(* IEC 61131-3 sources: codesys-api/examples/mqtt_large_payload/st/sfw, 5 files *)

(* ---- FB_MixedPushStream.st ---- *)
FUNCTION_BLOCK FB_MixedPushStream
// One periodic stream of the mixed-rate test through MQTT.MqttStoreForward (MixedPushTest, mixed_rate_test.py --push).
// FB_MixedStream's messages, built the same way (same tags, values, "MIX:<StreamId>:<round>:<part>:<parts>:<UTC ms>"
// header and "<tag>:<value>" lines, all parts back to back in Data), but each part is handed to the shared block Sfw
// with Push (a copy, so Data is rebuilt next round while earlier rounds are still held) instead of MQTTPublish blocks.
// QoS 1 only. The statistics keep FB_MixedStream's names and units, with these differences:
// - a period is never skipped because the previous round is still in flight: the block buffers it. Skipped counts
//   only periods a late scan jumped over; SkippedOffline the periods due while the broker was down (unless IsPushOffline);
// - TimeoutCount counts parts Push refused (not configured, AcceptPush FALSE, too large for a slot); drops and broker
//   refusals are the shared block's (MixedPushTest.DroppedCount, RefusedCount), not attributable to a stream;
// - a round is done when the block no longer holds anything pushed before or with it (ServiceRounds); send times run
//   from the build's end to that scan, so SendScans is at least 1; PartsDone counts the parts pushed in done rounds.
// Up to MAX_TRACKED rounds are timed at once; beyond that the oldest is forgotten (UntrackedCount, not in RoundsDone).
VAR CONSTANT
	MAX_BYTES : UDINT := 32000;
	MAX_PARTS : UINT := 64;
	MAX_TRACKED : UINT := 128;
	BOOL_COUNT : UINT := 1000;
	INT_COUNT : UINT := 500;
	REAL_COUNT : UINT := 500;
	MIN_PERIOD_US : ULINT := 10000;
END_VAR
VAR_INPUT
	IsEnabled : BOOL;
	StreamId : STRING(1);
	FirstTag : UINT;                        // 1 .. 2000, ScaleTest numbering: BOOL 1-1000, DINT 1001-1500, REAL 1501-2000
	LastTag : UINT;
	TagsPerMessage : UINT;
	Period : TIME;
	Topic : STRING(64);
	ToleranceUs : ULINT;                    // a period is due this much early (task jitter)
	IsPushOffline : BOOL;                   // push while the broker is down (the block holds it); FALSE skips, as FB_MixedStream
	BlockNowMs : UDINT;                     // SysTimeGetMs() taken just before the block's last call (MixedPushTest)
	ResetStats : BOOL;
END_VAR
VAR_IN_OUT
	Sfw : MQTT.MqttStoreForward;            // shared by both streams, owned and called by MixedPushTest
END_VAR
VAR_OUTPUT
	IsRoundActive : BOOL;                   // a pushed round still has a part in the block
END_VAR
VAR
	// Results, read online (microseconds unless named *Scans/*Count)
	Round : UDINT;                          // rounds started since download (not reset; the broker check uses it)
	RoundsStarted : UDINT;
	RoundsDone : UDINT;
	Skipped : UDINT;                        // periods a late scan jumped over (never for a round in flight)
	SkippedOffline : UDINT;                 // periods lost because the broker was not connected (IsPushOffline FALSE)
	PartsDone : UDINT;                      // parts pushed in the rounds that are done
	TimeoutCount : UDINT;                   // parts Push refused
	OverflowCount : UDINT;                  // rounds that did not fit MAX_BYTES / MAX_PARTS (not sent)
	LastBytes : UDINT;                      // all parts of the last round, headers included
	LastParts : UINT;
	LastBuildUs : UDINT;                    // value update + formatting of the whole round, in its first scan
	MaxBuildUs : UDINT;
	SumBuildUs : ULINT;
	LastSendUs : UDINT;                     // build finished -> the block holds nothing of the round (PUBACKs)
	MaxSendUs : UDINT;
	SumSendUs : ULINT;
	LastSendScans : UDINT;                  // scans from the build to that scan (at least 1)
	MaxSendScans : UDINT;
	SumSendScans : ULINT;
	MaxLateUs : UDINT;                      // how late after its due time a round started (scan phase)
	LastPushUs : UDINT;                     // the round's Push calls (copies into the block's storage)
	MaxPushUs : UDINT;
	SumPushUs : ULINT;
	MaxRoundsActive : UINT;                 // most rounds held at once
	UntrackedCount : UDINT;                 // rounds whose completion was not timed (more than MAX_TRACKED held)

	// State
	PartStart : ARRAY[0..MAX_PARTS - 1] OF UDINT;
	PartLength : ARRAY[0..MAX_PARTS - 1] OF UDINT;
	Data : ARRAY[0..MAX_BYTES - 1] OF BYTE;
	Bools : ARRAY[1..BOOL_COUNT] OF BOOL;
	Ints : ARRAY[1..INT_COUNT] OF DINT;
	Reals : ARRAY[1..REAL_COUNT] OF REAL;
	// rounds pushed and not yet done, oldest at TrackHead (a ring)
	TrackRequestUs : ARRAY[0..MAX_TRACKED - 1] OF ULINT;
	TrackPushMs : ARRAY[0..MAX_TRACKED - 1] OF UDINT;	// SysTimeGetMs() after the round's last Push
	TrackScan : ARRAY[0..MAX_TRACKED - 1] OF UDINT;
	TrackParts : ARRAY[0..MAX_TRACKED - 1] OF UINT;
	TrackHead : UINT;
	TrackCount : UINT;
	IsScheduled : BOOL;
	IsDue : BOOL;
	IsBuildOk : BOOL;
	NowTimeUs : ULINT;
	PeriodUs : ULINT;
	NextDueUs : ULINT;
	DueUs : ULINT;
	StepStartUs : ULINT;
	RequestUs : ULINT;
	ServiceNowUs : ULINT;
	ScanCount : UDINT;
	RoundParts : UINT;
	RoundPushed : UINT;
	Used : UDINT;
	Part : UINT;
	PartFirst : UINT;
	PartLast : UINT;
	Tag : UINT;
	Index : UINT;
	Kind : UDINT;
	StampMs : ULINT;
	StampText : STRING(24);
	Header : STRING(80);
	ValueText : STRING(40);
	RealValue : REAL;
END_VAR
// ---- implementation ----
ScanCount := ScanCount + 1;
IF ResetStats THEN
	RoundsStarted := 0; RoundsDone := 0; Skipped := 0; SkippedOffline := 0; PartsDone := 0; TimeoutCount := 0;
	OverflowCount := 0; MaxBuildUs := 0; SumBuildUs := 0; MaxSendUs := 0; SumSendUs := 0; MaxSendScans := 0;
	SumSendScans := 0; MaxLateUs := 0; MaxPushUs := 0; SumPushUs := 0; MaxRoundsActive := 0; UntrackedCount := 0;
END_IF

// What left the block since the last scan
ServiceRounds();

// Schedule: one round per Period, on a fixed grid from the scan that enabled the stream
NowTimeUs := NowUs();
PeriodUs := TIME_TO_ULINT(Period) * 1000;
IF NOT IsEnabled OR PeriodUs < MIN_PERIOD_US THEN
	IsScheduled := FALSE;
ELSIF NOT IsScheduled THEN
	IsScheduled := TRUE;
	NextDueUs := NowTimeUs;
END_IF
IsDue := FALSE;
IF IsScheduled AND NowTimeUs + ToleranceUs >= NextDueUs THEN
	IsDue := TRUE;
	DueUs := NextDueUs;
	NextDueUs := NextDueUs + PeriodUs;
	// a scan so late that whole periods passed: those are lost as well
	WHILE NowTimeUs + ToleranceUs >= NextDueUs DO
		NextDueUs := NextDueUs + PeriodUs;
		Skipped := Skipped + 1;
	END_WHILE
END_IF

IF IsDue THEN
	IF NOT PLC_PRG.IsBrokerConnected AND NOT IsPushOffline THEN
		SkippedOffline := SkippedOffline + 1;
	ELSIF FirstTag >= 1 AND LastTag >= FirstTag AND LastTag <= BOOL_COUNT + INT_COUNT + REAL_COUNT
		AND TagsPerMessage >= 1 THEN
		Round := Round + 1;
		RoundsStarted := RoundsStarted + 1;
		IF NowTimeUs > DueUs THEN
			MaxLateUs := MAX(MaxLateUs, ULINT_TO_UDINT(NowTimeUs - DueUs));
		END_IF
		StepStartUs := NowUs();
		// New values for this stream's tags: ScaleTest.UpdateValues' formulas with Round for Sequence
		FOR Tag := FirstTag TO LastTag DO
			IF Tag <= BOOL_COUNT THEN
				Bools[Tag] := ((UINT_TO_UDINT(Tag) + Round) MOD 3) = 0;
			ELSIF Tag <= BOOL_COUNT + INT_COUNT THEN
				Kind := UINT_TO_UDINT(Tag - BOOL_COUNT);
				Ints[Kind] := UDINT_TO_DINT((Kind * 37 + Round) MOD 20000) - 10000;
			ELSE
				Kind := UINT_TO_UDINT(Tag - BOOL_COUNT - INT_COUNT);
				Reals[Kind] := DINT_TO_REAL(UDINT_TO_DINT((Kind * 1237 + Round * 17) MOD 200000) - 100000) / 100.0;
			END_IF
		END_FOR
		SysTimeRtc.SysTimeRtcHighResGet(pTimestamp := StampMs);
		StampMs := LINT_TO_ULINT(ULINT_TO_LINT(StampMs) + ClockSync.OffsetMs);   // UTC, see ClockSync
		StampText := ULINT_TO_STRING(StampMs);

		// Every part of the round, back to back in Data (as FB_MixedStream)
		RoundParts := (LastTag - FirstTag + TagsPerMessage) / TagsPerMessage;
		IsBuildOk := RoundParts <= MAX_PARTS;
		Used := 0;
		PartFirst := FirstTag;
		Part := 0;
		WHILE IsBuildOk AND Part < RoundParts DO
			PartStart[Part] := Used;
			Header := CONCAT(CONCAT(CONCAT('MIX:', StreamId), ':'), UDINT_TO_STRING(Round));
			Header := CONCAT(CONCAT(CONCAT(Header, ':'), UINT_TO_STRING(Part)), ':');
			Header := CONCAT(CONCAT(CONCAT(CONCAT(Header, UINT_TO_STRING(RoundParts)), ':'), StampText), '$N');
			IsBuildOk := AppendZ(pBuffer := ADR(Data), Capacity := SIZEOF(Data), pText := ADR(Header), Used := Used);
			PartLast := MIN(LastTag, PartFirst + TagsPerMessage - 1);
			Tag := PartFirst;
			WHILE IsBuildOk AND Tag <= PartLast DO
				// formatted as ScaleTest.BuildTag formats each type
				IF Tag <= BOOL_COUNT THEN
					ValueText := SEL(Bools[Tag], '0', '1');
				ELSIF Tag <= BOOL_COUNT + INT_COUNT THEN
					ValueText := DINT_TO_STRING(Ints[Tag - BOOL_COUNT]);
				ELSE
					RealValue := Reals[Tag - BOOL_COUNT - INT_COUNT];
					ValueText := REAL_TO_STRING(DINT_TO_REAL(TRUNC(RealValue * 100.0 + SEL(RealValue >= 0.0, -0.5, 0.5))) / 100.0);
				END_IF
				IsBuildOk := AppendZ(pBuffer := ADR(Data), Capacity := SIZEOF(Data), pText := ADR(ScaleTest.Names[Tag]), Used := Used)
					AND_THEN AppendZ(pBuffer := ADR(Data), Capacity := SIZEOF(Data), pText := ADR(':'), Used := Used)
					AND_THEN AppendZ(pBuffer := ADR(Data), Capacity := SIZEOF(Data), pText := ADR(ValueText), Used := Used)
					AND_THEN AppendZ(pBuffer := ADR(Data), Capacity := SIZEOF(Data), pText := ADR('$N'), Used := Used);
				Tag := Tag + 1;
			END_WHILE
			PartLength[Part] := Used - PartStart[Part];
			PartFirst := PartLast + 1;
			Part := Part + 1;
		END_WHILE
		LastBuildUs := ULINT_TO_UDINT(NowUs() - StepStartUs);
		MaxBuildUs := MAX(MaxBuildUs, LastBuildUs);
		SumBuildUs := SumBuildUs + LastBuildUs;
		LastBytes := Used;
		LastParts := RoundParts;
		IF IsBuildOk THEN
			// Every part to the block, in order; the block hands them to the client in its call after both streams
			RequestUs := NowUs();
			RoundPushed := 0;
			FOR Part := 0 TO RoundParts - 1 DO
				IF Sfw.Push(Topic := ADR(Topic), Payload := ADR(Data[PartStart[Part]]), Length := PartLength[Part]) THEN
					RoundPushed := RoundPushed + 1;
				ELSE
					TimeoutCount := TimeoutCount + 1;
				END_IF
			END_FOR
			LastPushUs := ULINT_TO_UDINT(NowUs() - RequestUs);
			MaxPushUs := MAX(MaxPushUs, LastPushUs);
			SumPushUs := SumPushUs + LastPushUs;
			IF TrackCount >= MAX_TRACKED THEN
				// the oldest round is no longer timed; the newest still is, so IsRoundActive stays right
				TrackHead := (TrackHead + 1) MOD MAX_TRACKED;
				TrackCount := TrackCount - 1;
				UntrackedCount := UntrackedCount + 1;
			END_IF
			Index := (TrackHead + TrackCount) MOD MAX_TRACKED;
			TrackRequestUs[Index] := RequestUs;
			TrackPushMs[Index] := SysTimeCore.SysTimeGetMs();	// not before any part's push time in the block
			TrackScan[Index] := ScanCount;
			TrackParts[Index] := RoundPushed;
			TrackCount := TrackCount + 1;
			MaxRoundsActive := MAX(MaxRoundsActive, TrackCount);
			IsRoundActive := TRUE;
			// no ServiceRounds here: the block's outputs are fresh only after its call, later in this scan
		ELSE
			OverflowCount := OverflowCount + 1;
		END_IF
	END_IF
END_IF

(* ---- MixedPushTest.st ---- *)
PROGRAM MixedPushTest
// MixedTest's mixed-rate load through MQTT.MqttStoreForward (library 1.4.0.0) instead of MQTTPublish pools: the same
// two streams, messages and statistics (FB_MixedPushStream), each message handed to the block with Push. QoS 1 only.
// mixed_rate_test.py --push drives it. Called by PLC_PRG after StoreForwardTest, before the end-of-scan client call;
// PLC_PRG makes that call when IsLiveHandedOff, and CallClient keeps calling while IsSendInFlight, early stop on
// IsUnsentPending while IsEnabled (patch_demo_store_forward.py adds all three, in the MQTT 5 demo copy only).
// One block for both streams, as a comms program would have it: one buffer, one call per scan after both streams'
// pushes, one set of lanes and out slots, one live-first fence. Scan figures are PLC_PRG's of the scan before.
VAR CONSTANT
	LINE_BYTES : UDINT := 24;               // a "<tag>:<value>" line, worst case with margin (9-char name, measured mean 13-16 B)
	HEADER_BYTES : UDINT := 64;             // "MIX:..." header line, with room to spare
	MAX_SLOT_BYTES : UDINT := 32000;        // FB_MixedPushStream.MAX_BYTES: no part is larger than a round
END_VAR
VAR
	// Settings, written online
	IsEnabled : BOOL;                       // configures the block on the first enable
	SlowTagsPerMessage : UINT := 1500;
	FastTagsPerMessage : UINT := 500;
	SlowPeriod : TIME := T#1S;
	FastPeriod : TIME := T#100MS;
	ToleranceUs : ULINT := 20000;
	IsPushOffline : BOOL;                   // push while the broker is down (held); FALSE skips those periods, as MixedTest
	ResetStats : BOOL;
	// the block's configuration: on the first enable and on ConfigureRequest (with the block idle: Reset refuses while
	// a sample is in the client, and the configuration is then retried every scan while IsEnabled)
	LiveLanes : UINT := 2;
	BacklogLanes : UINT := 4;
	SlotTopicSize : UINT := 64;
	SlotPayloadSize : UDINT := 0;           // 0: from the larger TagsPerMessage, LINE_BYTES a tag + HEADER_BYTES (<= MAX_SLOT_BYTES)
	StorageBytes : UDINT := 262144;         // part of Storage given to Configure
	ConfigureRequest : BOOL;                // Reset(Discard) and Configure again with the settings above
	// the block's runtime inputs, passed every call
	BacklogStartsPerCall : UINT := 2;
	BacklogBytesPerCall : UDINT := 8192;
	ReservedOutSlots : UINT := 2;
	ReservedCredits : UINT := 2;
	IsHoldOnNoSubscribers : BOOL := TRUE;
	NoSubscriberPause : TIME := T#5S;

	Slow : FB_MixedPushStream;
	Fast : FB_MixedPushStream;
	Sfw : MQTT.MqttStoreForward;
	Storage : ARRAY[0..262143] OF BYTE;       // 256 KiB, keeps the application small (RealisticSfwTest has the big buffer)
	IsSendInFlight : BOOL;                  // PLC_PRG.CallClient keeps calling the client while this is TRUE
	IsLiveHandedOff : BOOL;                 // PLC_PRG makes the end-of-scan client call
	BlockNowMs : UDINT;                     // SysTimeGetMs() just before the block's call, for the streams' next scan
	SlotBytes : UDINT;
	StartUs : ULINT;

	// Results, read online
	ScanCount : UDINT;                      // scans while enabled
	SumCycleUs : ULINT;
	MaxCycleUs : UDINT;
	SumScanClientUs : ULINT;
	MaxScanClientUs : UDINT;
	MaxIntervalUs : UDINT;
	MinIntervalUs : UDINT := 16#FFFFFFFF;
	SumClientCalls : ULINT;
	IsCounting : BOOL;
	IsConfigured : BOOL;
	ConfigureCount : UDINT;
	ConfiguredSlotBytes : UDINT;
	LastConfigureError : MQTT.STORE_FORWARD_ERROR;
	Capacity : UINT;                        // slots
	// the block's counters since download (mixed_rate_test.py takes differences)
	PushedCount : ULINT;
	DeliveredCount : ULINT;
	DroppedCount : ULINT;
	RefusedCount : ULINT;
	DiscardedCount : ULINT;
	LiveDeferredCount : ULINT;
	NotAcceptedCount : ULINT;
	InvalidCount : ULINT;
	// the block's state after its call, and maxima since ResetStats
	QueuedCount : UINT;
	InFlightCount : UINT;
	HasWork : BOOL;
	MaxQueuedCount : UINT;
	MaxInFlightCount : UINT;
	MaxOldestAgeMs : UDINT;
	BlockUs : UDINT;                        // the block's call, every scan
	MaxBlockUs : UDINT;
	SumBlockUs : ULINT;                     // while IsEnabled (over ScanCount)
	LiveHandOffScans : UDINT;
END_VAR
// ---- implementation ----
IF ResetStats THEN
	ScanCount := 0; SumCycleUs := 0; MaxCycleUs := 0; SumScanClientUs := 0; MaxScanClientUs := 0;
	MaxIntervalUs := 0; MinIntervalUs := 16#FFFFFFFF; SumClientCalls := 0;
	MaxQueuedCount := 0; MaxInFlightCount := 0; MaxOldestAgeMs := 0; MaxBlockUs := 0; SumBlockUs := 0;
	LiveHandOffScans := 0;
END_IF
IF IsCounting THEN
	ScanCount := ScanCount + 1;
	SumCycleUs := SumCycleUs + PLC_PRG.CycleUs;
	MaxCycleUs := MAX(MaxCycleUs, PLC_PRG.CycleUs);
	SumScanClientUs := SumScanClientUs + PLC_PRG.ScanClientUs;
	MaxScanClientUs := MAX(MaxScanClientUs, PLC_PRG.ScanClientUs);
	MaxIntervalUs := MAX(MaxIntervalUs, PLC_PRG.IntervalUs);
	MinIntervalUs := MIN(MinIntervalUs, PLC_PRG.IntervalUs);
	SumClientCalls := SumClientCalls + INT_TO_ULINT(PLC_PRG.ClientCall);
END_IF
IsCounting := IsEnabled;

// Configure before the first push (after SetMqttInOut: Configure reads COM_CONFIG.CountSlotsOut)
IF ConfigureRequest OR (IsEnabled AND NOT IsConfigured) THEN
	ConfigureRequest := FALSE;
	SlotBytes := SlotPayloadSize;
	IF SlotBytes = 0 THEN
		SlotBytes := MIN(MAX_SLOT_BYTES,
			UINT_TO_UDINT(MAX(SlowTagsPerMessage, FastTagsPerMessage)) * LINE_BYTES + HEADER_BYTES);
	END_IF
	Sfw.Reset(Discard := TRUE);
	Sfw.SetMqttInOut(MQTT_IN_OUT := PLC_PRG.MqttLink);
	IsConfigured := Sfw.Configure(Storage := ADR(Storage), StorageSize := MIN(StorageBytes, SIZEOF(Storage)),
		SlotTopicSize := SlotTopicSize, SlotPayloadSize := SlotBytes, LiveLanes := LiveLanes,
		BacklogLanes := BacklogLanes);
	ConfigureCount := ConfigureCount + 1;
	ConfiguredSlotBytes := SlotBytes;
	LastConfigureError := Sfw.LastConfigureError;
END_IF

Slow(IsEnabled := IsEnabled, StreamId := 'S', FirstTag := 1, LastTag := 1500, TagsPerMessage := SlowTagsPerMessage,
	Period := SlowPeriod, Topic := 'raw_data_demo/mixed/slow', ToleranceUs := ToleranceUs,
	IsPushOffline := IsPushOffline, BlockNowMs := BlockNowMs, ResetStats := ResetStats, Sfw := Sfw);
Fast(IsEnabled := IsEnabled, StreamId := 'F', FirstTag := 1501, LastTag := 2000, TagsPerMessage := FastTagsPerMessage,
	Period := FastPeriod, Topic := 'raw_data_demo/mixed/fast', ToleranceUs := ToleranceUs,
	IsPushOffline := IsPushOffline, BlockNowMs := BlockNowMs, ResetStats := ResetStats, Sfw := Sfw);
ResetStats := FALSE;

// Once per scan, after both streams' pushes: this scan's samples to the client, then backlog if admitted
BlockNowMs := SysTimeCore.SysTimeGetMs();
StartUs := NowUs();
Sfw(AcceptPush := TRUE, Enable := TRUE, IsHoldOnNoSubscribers := IsHoldOnNoSubscribers,
	NoSubscriberPause := NoSubscriberPause, BacklogStartsPerCall := BacklogStartsPerCall,
	BacklogBytesPerCall := BacklogBytesPerCall, ReservedOutSlots := ReservedOutSlots, ReservedCredits := ReservedCredits,
	IsInferRefusals := FALSE);
BlockUs := ULINT_TO_UDINT(NowUs() - StartUs);
MaxBlockUs := MAX(MaxBlockUs, BlockUs);
IF IsEnabled THEN
	SumBlockUs := SumBlockUs + BlockUs;
END_IF

Capacity := Sfw.Capacity;
PushedCount := Sfw.PushedCount;
DeliveredCount := Sfw.DeliveredCount;
DroppedCount := Sfw.DroppedCount;
RefusedCount := Sfw.RefusedCount + Sfw.InferredRefusedCount;
DiscardedCount := Sfw.DiscardedCount;
LiveDeferredCount := Sfw.LiveDeferredCount;
NotAcceptedCount := Sfw.NotAcceptedCount;
InvalidCount := Sfw.InvalidCount;
QueuedCount := Sfw.QueuedCount;
InFlightCount := Sfw.InFlightCount;
HasWork := Sfw.HasWork;
MaxQueuedCount := MAX(MaxQueuedCount, QueuedCount);
MaxInFlightCount := MAX(MaxInFlightCount, InFlightCount);
MaxOldestAgeMs := MAX(MaxOldestAgeMs, Sfw.OldestAgeMs);
IsSendInFlight := Sfw.InFlightCount > 0;
IsLiveHandedOff := Sfw.IsLiveHandedOff;
IF IsLiveHandedOff THEN
	LiveHandOffScans := LiveHandOffScans + 1;
END_IF

(* ---- RealisticSfwTest.BuildPayload.st ---- *)
// Action BuildPayload: Payload := _TS:<BuildStampMs>, <BuildSeqKey><BuildSeq>, then padding lines p:000... of at most
// PAD_LINE_CHARS characters until Used is within 3 bytes of BuildTargetBytes (or of the end of Payload). Used is the
// payload's length. Direct byte writes: CONCAT stops at 255 characters.
// ---- implementation ----
Used := 0;
AppendText(pBuffer := ADR(Payload), Capacity := SIZEOF(Payload), Text := CONCAT('_TS:', ULINT_TO_STRING(BuildStampMs)),
	Used := Used);
AppendText(pBuffer := ADR(Payload), Capacity := SIZEOF(Payload),
	Text := CONCAT(CONCAT('$L', BuildSeqKey), UDINT_TO_STRING(BuildSeq)), Used := Used);
PayloadLimit := MIN(BuildTargetBytes, SIZEOF(Payload) - 1);
pPayload := ADR(Payload);
// a padding line is a line feed, 'p:' and at least one '0'; stop when less than that is left
WHILE Used + 4 <= PayloadLimit DO
	LineChars := MIN(PayloadLimit - Used - 1, PAD_LINE_CHARS);
	pPayload[Used] := 16#0A;	// line feed
	pPayload[Used + 1] := 16#70;	// 'p'
	pPayload[Used + 2] := 16#3A;	// ':'
	Used := Used + 3;
	FOR PadIndex := 3 TO LineChars DO
		pPayload[Used] := 16#30;	// '0'
		Used := Used + 1;
	END_FOR
END_WHILE
pPayload[Used] := 0;

(* ---- RealisticSfwTest.st ---- *)
PROGRAM RealisticSfwTest
// A realistic two-stream outage load through MQTT.MqttStoreForward (library 1.4.0.0, or the adaptive version with the
// same Configure): Slow pushes one ~SlowBytes sample per SlowPeriod on SlowTopic, Fast one ~FastBytes sample per
// FastPeriod on FastTopic, each stamped with the PLC's UTC time when captured. sfw_test.py realistic drives it.
// Payload, "lines" for Marigraf: _TS:<UTC ms>, sfw_slow_seq:<n> or sfw_fast_seq:<n>, then p:000... padding lines of at
// most PAD_LINE_CHARS characters (Marigraf drops lines over 4,096 bytes) up to the target size (BuildPayload).
// IsTwoBlocks: BlockSlow and BlockFast, each with its own slot size and its share of Storage (StorageShareSlowPercent);
// FALSE: BlockSlow takes both streams over all of StorageBytes, its slots sized for the larger sample. The mode is
// latched by the configuration (IsTwoBlocksConfigured); change it with ConfigureRequest.
// Called by PLC_PRG after MixedPushTest, before the end-of-scan client call; PLC_PRG makes that call when
// IsLiveHandedOff, and CallClient keeps calling while IsSendInFlight, early stop on IsUnsentPending while IsEnabled
// (patch_demo_store_forward.py adds all three, in the MQTT 5 demo copy only).
VAR CONSTANT
	PAD_LINE_CHARS : UDINT := 100;          // a padding line "p:000...", line feed not counted
	SLOT_ROUND_BYTES : UDINT := 1024;       // a slot size of 0 is the sample size rounded up to this
	STORAGE_ALIGN : UDINT := 8;             // BlockFast's share starts on this boundary
END_VAR
VAR
	// Settings, written online
	IsEnabled : BOOL;                       // configures on the first enable, then pushes both streams
	IsPushing : BOOL := TRUE;               // FALSE: keep calling the blocks (drain) without new samples
	SlowPeriod : TIME := T#1S;
	SlowBytes : UDINT := 26000;             // payload size, about (padding lines stop within 3 bytes of it)
	SlowTopic : STRING(64) := 'raw_data/sfw/slow';
	FastPeriod : TIME := T#100MS;
	FastBytes : UDINT := 5000;
	FastTopic : STRING(64) := 'raw_data/sfw/fast';
	ResetStats : BOOL;
	// the configuration: on the first enable and on ConfigureRequest (Reset(Discard) first; Reset and Configure refuse
	// while a sample is in the client, and the configuration is then retried every scan while IsEnabled)
	IsTwoBlocks : BOOL := TRUE;
	StorageBytes : UDINT := 2621440;        // part of Storage given to the block(s)
	StorageShareSlowPercent : UDINT := 33;  // two blocks: BlockSlow's share of StorageBytes, BlockFast has the rest
	SlotTopicSize : UINT := 64;
	SlowSlotPayloadSize : UDINT := 0;       // 0: SlowBytes rounded up to SLOT_ROUND_BYTES
	FastSlotPayloadSize : UDINT := 0;       // 0: FastBytes rounded up; one block: the larger of the two slot sizes
	SlowLiveLanes : UINT := 1;              // two blocks
	SlowBacklogLanes : UINT := 2;
	FastLiveLanes : UINT := 1;
	FastBacklogLanes : UINT := 2;
	OneBlockLiveLanes : UINT := 2;          // one block
	OneBlockBacklogLanes : UINT := 4;
	ConfigureRequest : BOOL;                // Reset(Discard) and Configure again with the settings above
	// the blocks' runtime inputs, passed to both every call
	BacklogStartsPerCall : UINT := 3;
	BacklogBytesPerCall : UDINT := 16383;
	ReservedOutSlots : UINT := 2;
	ReservedCredits : UINT := 2;
	IsHoldOnNoSubscribers : BOOL := TRUE;
	NoSubscriberPause : TIME := T#5S;

	BlockSlow : MQTT.MqttStoreForward;
	BlockFast : MQTT.MqttStoreForward;      // idle (not configured) with one block
	Storage : ARRAY[0..2621439] OF BYTE;      // 2.5 MiB, one array for both blocks (the P2CDS-622 refused larger buffers)
	Payload : STRING(32767);
	pStorage : POINTER TO BYTE;
	TotalBytes : UDINT;
	IsSlowConfigured : BOOL;
	IsFastConfigured : BOOL;
	IsSlowDue : BOOL;
	IsFastDue : BOOL;
	NowPushUs : ULINT;
	PeriodUs : ULINT;
	NextSlowUs : ULINT;
	NextFastUs : ULINT;
	StampMs : ULINT;
	LastSlowStampMs : ULINT;
	LastFastStampMs : ULINT;
	IsPushed : BOOL;
	StartUs : ULINT;
	// BuildPayload's inputs and work
	BuildStampMs : ULINT;
	BuildSeqKey : STRING(16);               // 'sfw_slow_seq:' or 'sfw_fast_seq:'
	BuildSeq : UDINT;
	BuildTargetBytes : UDINT;
	Used : UDINT;                           // BuildPayload's result: the payload's length
	pPayload : POINTER TO BYTE;
	PayloadLimit : UDINT;
	LineChars : UDINT;
	PadIndex : UDINT;

	// Results, read online (the blocks' own outputs: BlockSlow.<output>, BlockFast.<output>)
	IsConfigured : BOOL;
	IsTwoBlocksConfigured : BOOL;
	ConfigureCount : UDINT;
	SlowSlotBytes : UDINT;                  // the configured slot payload sizes and storage shares
	FastSlotBytes : UDINT;
	SlowStorageBytes : UDINT;
	FastStorageBytes : UDINT;
	LastSlowConfigureError : MQTT.STORE_FORWARD_ERROR;
	LastFastConfigureError : MQTT.STORE_FORWARD_ERROR;
	SlowNextSeq : UDINT;                    // the sequence of the next sample (the first is 1)
	FastNextSeq : UDINT;
	SlowPushFailCount : UDINT;
	FastPushFailCount : UDINT;
	SlowSkippedCount : UDINT;               // periods skipped by a resynchronisation (a scan more than a period late)
	FastSkippedCount : UDINT;
	SlowPushUs : UDINT;                     // building the payload and the Push
	MaxSlowPushUs : UDINT;
	FastPushUs : UDINT;
	MaxFastPushUs : UDINT;
	SlowBlockUs : UDINT;                    // the block's call, every scan
	MaxSlowBlockUs : UDINT;
	FastBlockUs : UDINT;
	MaxFastBlockUs : UDINT;
	HasWork : BOOL;                         // either block holds a sample
	IsSendInFlight : BOOL;                  // PLC_PRG.CallClient keeps calling the client while this is TRUE
	IsLiveHandedOff : BOOL;                 // PLC_PRG makes the end-of-scan client call
	LiveHandOffScans : UDINT;
END_VAR
// ---- implementation ----
IF ResetStats THEN
	ResetStats := FALSE;
	SlowPushFailCount := 0; FastPushFailCount := 0; SlowSkippedCount := 0; FastSkippedCount := 0;
	MaxSlowPushUs := 0; MaxFastPushUs := 0; MaxSlowBlockUs := 0; MaxFastBlockUs := 0; LiveHandOffScans := 0;
END_IF

// Configure before the first push (after SetMqttInOut: Configure reads COM_CONFIG.CountSlotsOut)
IF ConfigureRequest OR (IsEnabled AND NOT IsConfigured) THEN
	ConfigureRequest := FALSE;
	IsTwoBlocksConfigured := IsTwoBlocks;
	TotalBytes := MIN(StorageBytes, SIZEOF(Storage));
	SlowSlotBytes := SlowSlotPayloadSize;
	IF SlowSlotBytes = 0 THEN
		SlowSlotBytes := (SlowBytes + SLOT_ROUND_BYTES - 1) / SLOT_ROUND_BYTES * SLOT_ROUND_BYTES;
	END_IF
	FastSlotBytes := FastSlotPayloadSize;
	IF FastSlotBytes = 0 THEN
		FastSlotBytes := (FastBytes + SLOT_ROUND_BYTES - 1) / SLOT_ROUND_BYTES * SLOT_ROUND_BYTES;
	END_IF
	IF IsTwoBlocksConfigured THEN
		SlowStorageBytes := TotalBytes * MIN(StorageShareSlowPercent, 100) / 100 / STORAGE_ALIGN * STORAGE_ALIGN;
		FastStorageBytes := TotalBytes - SlowStorageBytes;
	ELSE
		SlowSlotBytes := MAX(SlowSlotBytes, FastSlotBytes);
		FastSlotBytes := 0;
		SlowStorageBytes := TotalBytes;
		FastStorageBytes := 0;
	END_IF
	BlockSlow.Reset(Discard := TRUE);
	BlockFast.Reset(Discard := TRUE);
	BlockSlow.SetMqttInOut(MQTT_IN_OUT := PLC_PRG.MqttLink);
	BlockFast.SetMqttInOut(MQTT_IN_OUT := PLC_PRG.MqttLink);
	pStorage := ADR(Storage);
	IF IsTwoBlocksConfigured THEN
		IsSlowConfigured := BlockSlow.Configure(Storage := pStorage, StorageSize := SlowStorageBytes,
			SlotTopicSize := SlotTopicSize, SlotPayloadSize := SlowSlotBytes, LiveLanes := SlowLiveLanes,
			BacklogLanes := SlowBacklogLanes);
		IsFastConfigured := BlockFast.Configure(Storage := pStorage + SlowStorageBytes, StorageSize := FastStorageBytes,
			SlotTopicSize := SlotTopicSize, SlotPayloadSize := FastSlotBytes, LiveLanes := FastLiveLanes,
			BacklogLanes := FastBacklogLanes);
	ELSE
		IsSlowConfigured := BlockSlow.Configure(Storage := pStorage, StorageSize := SlowStorageBytes,
			SlotTopicSize := SlotTopicSize, SlotPayloadSize := SlowSlotBytes, LiveLanes := OneBlockLiveLanes,
			BacklogLanes := OneBlockBacklogLanes);
		IsFastConfigured := TRUE;
	END_IF
	IsConfigured := IsSlowConfigured AND IsFastConfigured;
	ConfigureCount := ConfigureCount + 1;
	LastSlowConfigureError := BlockSlow.LastConfigureError;
	LastFastConfigureError := BlockFast.LastConfigureError;
	IF SlowNextSeq = 0 THEN
		SlowNextSeq := 1;
	END_IF
	IF FastNextSeq = 0 THEN
		FastNextSeq := 1;
	END_IF
END_IF

// fixed schedules (a TON restarted on its Q runs a scan or two slow per period); resynchronised after a pause
IsSlowDue := FALSE;
IsFastDue := FALSE;
IF IsEnabled AND IsPushing THEN
	NowPushUs := NowUs();
	PeriodUs := MAX(TIME_TO_ULINT(SlowPeriod), 1) * 1000;
	IF NextSlowUs = 0 OR NowPushUs > NextSlowUs + PeriodUs THEN
		IF NextSlowUs <> 0 THEN
			SlowSkippedCount := SlowSkippedCount + ULINT_TO_UDINT((NowPushUs - NextSlowUs) / PeriodUs);
		END_IF
		NextSlowUs := NowPushUs;
	END_IF
	IF NowPushUs >= NextSlowUs THEN
		IsSlowDue := TRUE;
		NextSlowUs := NextSlowUs + PeriodUs;
	END_IF
	PeriodUs := MAX(TIME_TO_ULINT(FastPeriod), 1) * 1000;
	IF NextFastUs = 0 OR NowPushUs > NextFastUs + PeriodUs THEN
		IF NextFastUs <> 0 THEN
			FastSkippedCount := FastSkippedCount + ULINT_TO_UDINT((NowPushUs - NextFastUs) / PeriodUs);
		END_IF
		NextFastUs := NowPushUs;
	END_IF
	IF NowPushUs >= NextFastUs THEN
		IsFastDue := TRUE;
		NextFastUs := NextFastUs + PeriodUs;
	END_IF
ELSE
	NextSlowUs := 0;
	NextFastUs := 0;
END_IF

IF IsSlowDue THEN
	StartUs := NowUs();
	// the capture time, unique and increasing per stream so Marigraf keeps every sample
	SysTimeRtc.SysTimeRtcHighResGet(pTimestamp := StampMs);
	IF StampMs <= LastSlowStampMs THEN
		StampMs := LastSlowStampMs + 1;
	END_IF
	LastSlowStampMs := StampMs;
	BuildStampMs := StampMs;
	BuildSeqKey := 'sfw_slow_seq:';
	BuildSeq := SlowNextSeq;
	BuildTargetBytes := SlowBytes;
	BuildPayload();
	IsPushed := BlockSlow.Push(Topic := ADR(SlowTopic), Payload := ADR(Payload), Length := Used);
	IF IsPushed THEN
		SlowNextSeq := SlowNextSeq + 1;
	ELSE
		SlowPushFailCount := SlowPushFailCount + 1;
	END_IF
	SlowPushUs := ULINT_TO_UDINT(NowUs() - StartUs);
	MaxSlowPushUs := MAX(MaxSlowPushUs, SlowPushUs);
END_IF

IF IsFastDue THEN
	StartUs := NowUs();
	SysTimeRtc.SysTimeRtcHighResGet(pTimestamp := StampMs);
	IF StampMs <= LastFastStampMs THEN
		StampMs := LastFastStampMs + 1;
	END_IF
	LastFastStampMs := StampMs;
	BuildStampMs := StampMs;
	BuildSeqKey := 'sfw_fast_seq:';
	BuildSeq := FastNextSeq;
	BuildTargetBytes := FastBytes;
	BuildPayload();
	IF IsTwoBlocksConfigured THEN
		IsPushed := BlockFast.Push(Topic := ADR(FastTopic), Payload := ADR(Payload), Length := Used);
	ELSE
		IsPushed := BlockSlow.Push(Topic := ADR(FastTopic), Payload := ADR(Payload), Length := Used);
	END_IF
	IF IsPushed THEN
		FastNextSeq := FastNextSeq + 1;
	ELSE
		FastPushFailCount := FastPushFailCount + 1;
	END_IF
	FastPushUs := ULINT_TO_UDINT(NowUs() - StartUs);
	MaxFastPushUs := MAX(MaxFastPushUs, FastPushUs);
END_IF

// Once per scan, after both streams' pushes: this scan's samples to the client, then backlog if admitted. BlockFast
// is called with one block too (not configured, it returns at once), so a mode change lets nothing hang.
StartUs := NowUs();
BlockSlow(AcceptPush := TRUE, Enable := TRUE, IsHoldOnNoSubscribers := IsHoldOnNoSubscribers,
	NoSubscriberPause := NoSubscriberPause, BacklogStartsPerCall := BacklogStartsPerCall,
	BacklogBytesPerCall := BacklogBytesPerCall, ReservedOutSlots := ReservedOutSlots, ReservedCredits := ReservedCredits,
	IsInferRefusals := FALSE);
SlowBlockUs := ULINT_TO_UDINT(NowUs() - StartUs);
MaxSlowBlockUs := MAX(MaxSlowBlockUs, SlowBlockUs);
StartUs := NowUs();
BlockFast(AcceptPush := TRUE, Enable := TRUE, IsHoldOnNoSubscribers := IsHoldOnNoSubscribers,
	NoSubscriberPause := NoSubscriberPause, BacklogStartsPerCall := BacklogStartsPerCall,
	BacklogBytesPerCall := BacklogBytesPerCall, ReservedOutSlots := ReservedOutSlots, ReservedCredits := ReservedCredits,
	IsInferRefusals := FALSE);
FastBlockUs := ULINT_TO_UDINT(NowUs() - StartUs);
MaxFastBlockUs := MAX(MaxFastBlockUs, FastBlockUs);

HasWork := BlockSlow.HasWork OR BlockFast.HasWork;
IsSendInFlight := BlockSlow.InFlightCount > 0 OR BlockFast.InFlightCount > 0;
IsLiveHandedOff := BlockSlow.IsLiveHandedOff OR BlockFast.IsLiveHandedOff;
IF IsLiveHandedOff THEN
	LiveHandOffScans := LiveHandOffScans + 1;
END_IF

(* ---- StoreForwardTest.st ---- *)
PROGRAM StoreForwardTest
// Store-and-forward test of MQTT.MqttStoreForward (library 1.4.0.0): sequence-numbered samples stamped with the
// PLC's UTC time when captured, on Topic, through the block on PLC_PRG.MqttLink. sfw_test.py drives it.
// Payload, "lines" for Marigraf: _TS:<UTC ms>, sfw_seq:<sequence>, and with PadBytes an sfw_pad line.
// Called by PLC_PRG after the publishers and before the end-of-scan client call; PLC_PRG makes that call when
// IsLiveHandedOff, and CallClient keeps calling while IsSendInFlight, early stop on IsUnsentPending.
VAR
	// Settings, written online
	IsEnabled : BOOL;                       // configures the block once, then pushes every PushPeriod
	IsPushing : BOOL := TRUE;               // FALSE: keep calling the block (drain) without new samples
	PushPeriod : TIME := T#100MS;
	PushesPerTick : UINT := 1;              // samples per tick, a burst within one scan
	PadBytes : UINT := 0;                   // extra payload bytes in an sfw_pad line
	Topic : STRING(64) := 'raw_data/sfw/bench';
	SlotTopicSize : UINT := 64;
	SlotPayloadSize : UDINT := 2048;
	LiveLanes : UINT := 2;
	BacklogLanes : UINT := 4;
	StorageBytes : UDINT := 262144;         // part of Storage given to Configure (a small value tests overflow)
	ConfigureRequest : BOOL;                // Reset(Discard) and Configure again with the settings above
	CheckRequest : BOOL;                    // CheckOwnership once
	IsCheckEveryScan : BOOL;                // CheckOwnership in every scan (costs a walk of every slot)
	ResetStats : BOOL;
	// the block's runtime inputs, passed every call
	Enable : BOOL := TRUE;
	AcceptPush : BOOL := TRUE;
	IsHoldOnNoSubscribers : BOOL := TRUE;
	NoSubscriberPause : TIME := T#5S;
	BacklogStartsPerCall : UINT := 2;
	BacklogBytesPerCall : UDINT := 8192;
	ReservedOutSlots : UINT := 2;
	ReservedCredits : UINT := 2;
	IsInferRefusals : BOOL;

	Telemetry : MQTT.MqttStoreForward;
	Storage : ARRAY[0..262143] OF BYTE;       // 256 KiB, keeps the application small (RealisticSfwTest has the big buffer)
	Payload : STRING(32767);
	IsPushDue : BOOL;
	NowPushUs : ULINT;
	NextPushUs : ULINT;
	PeriodUs : ULINT;
	StampMs : ULINT;
	LastStampMs : ULINT;
	Used : UDINT;
	pPayload : POINTER TO BYTE;
	PadIndex : UINT;
	Burst : UINT;
	StartUs : ULINT;

	// Results, read online
	IsConfigured : BOOL;
	ConfigureCount : UDINT;
	NextSequence : UDINT;                   // the sequence of the next sample (the first is 1)
	PushFailCount : UDINT;
	CheckCount : UDINT;
	CheckFailCount : UDINT;
	PushUs : UDINT;
	MaxPushUs : UDINT;
	BlockUs : UDINT;
	MaxBlockUs : UDINT;
	IsSendInFlight : BOOL;                  // PLC_PRG.CallClient keeps calling the client while this is TRUE
	IsLiveHandedOff : BOOL;                 // PLC_PRG makes the end-of-scan client call
	LiveHandOffScans : UDINT;
END_VAR
// ---- implementation ----
IF ResetStats THEN
	ResetStats := FALSE;
	PushFailCount := 0; CheckCount := 0; CheckFailCount := 0; MaxPushUs := 0; MaxBlockUs := 0; LiveHandOffScans := 0;
END_IF
IF ConfigureRequest OR (IsEnabled AND NOT IsConfigured) THEN
	ConfigureRequest := FALSE;
	Telemetry.Reset(Discard := TRUE);
	Telemetry.SetMqttInOut(MQTT_IN_OUT := PLC_PRG.MqttLink);
	IsConfigured := Telemetry.Configure(Storage := ADR(Storage), StorageSize := MIN(StorageBytes, SIZEOF(Storage)),
		SlotTopicSize := SlotTopicSize, SlotPayloadSize := SlotPayloadSize, LiveLanes := LiveLanes,
		BacklogLanes := BacklogLanes);
	ConfigureCount := ConfigureCount + 1;
	IF NextSequence = 0 THEN
		NextSequence := 1;
	END_IF
END_IF

// a fixed schedule (a TON restarted on its Q runs a scan or two slow per period); resynchronised after a pause
IsPushDue := FALSE;
IF IsEnabled AND IsPushing THEN
	NowPushUs := NowUs();
	PeriodUs := TIME_TO_ULINT(PushPeriod) * 1000;
	IF NextPushUs = 0 OR NowPushUs > NextPushUs + PeriodUs THEN
		NextPushUs := NowPushUs;
	END_IF
	IF NowPushUs >= NextPushUs THEN
		IsPushDue := TRUE;
		NextPushUs := NextPushUs + PeriodUs;
	END_IF
ELSE
	NextPushUs := 0;
END_IF
IF IsPushDue THEN
	FOR Burst := 1 TO MAX(PushesPerTick, 1) DO
		StartUs := NowUs();
		// the capture time, unique per sample so Marigraf keeps every one
		SysTimeRtc.SysTimeRtcHighResGet(pTimestamp := StampMs);
		IF StampMs <= LastStampMs THEN
			StampMs := LastStampMs + 1;
		END_IF
		LastStampMs := StampMs;
		Used := 0;
		AppendText(pBuffer := ADR(Payload), Capacity := SIZEOF(Payload), Text := CONCAT('_TS:', ULINT_TO_STRING(StampMs)), Used := Used);
		AppendText(pBuffer := ADR(Payload), Capacity := SIZEOF(Payload), Text := CONCAT('$Lsfw_seq:', UDINT_TO_STRING(NextSequence)), Used := Used);
		IF PadBytes > 0 THEN
			AppendText(pBuffer := ADR(Payload), Capacity := SIZEOF(Payload), Text := '$Lsfw_pad:', Used := Used);
			pPayload := ADR(Payload);
			FOR PadIndex := 1 TO PadBytes DO
				IF Used + 1 < SIZEOF(Payload) THEN
					pPayload[Used] := 16#30;	// '0'
					Used := Used + 1;
				END_IF
			END_FOR
			pPayload[Used] := 0;
		END_IF
		IF Telemetry.Push(Topic := ADR(Topic), Payload := ADR(Payload), Length := Used) THEN
			NextSequence := NextSequence + 1;
		ELSE
			PushFailCount := PushFailCount + 1;
		END_IF
		PushUs := ULINT_TO_UDINT(NowUs() - StartUs);
		MaxPushUs := MAX(MaxPushUs, PushUs);
	END_FOR
END_IF

StartUs := NowUs();
Telemetry(AcceptPush := AcceptPush, Enable := Enable, IsHoldOnNoSubscribers := IsHoldOnNoSubscribers,
	NoSubscriberPause := NoSubscriberPause, BacklogStartsPerCall := BacklogStartsPerCall,
	BacklogBytesPerCall := BacklogBytesPerCall, ReservedOutSlots := ReservedOutSlots, ReservedCredits := ReservedCredits,
	IsInferRefusals := IsInferRefusals);
BlockUs := ULINT_TO_UDINT(NowUs() - StartUs);
MaxBlockUs := MAX(MaxBlockUs, BlockUs);

IF CheckRequest OR IsCheckEveryScan THEN
	CheckRequest := FALSE;
	CheckCount := CheckCount + 1;
	IF NOT Telemetry.CheckOwnership() THEN
		CheckFailCount := CheckFailCount + 1;
	END_IF
END_IF
IsSendInFlight := Telemetry.InFlightCount > 0;
IsLiveHandedOff := Telemetry.IsLiveHandedOff;
IF IsLiveHandedOff THEN
	LiveHandOffScans := LiveHandOffScans + 1;
END_IF
